Fanuc KAREL source: KS00006.KL

PROGRAM KS00006
%NOLOCKGROUP
TYPE
  REC_T = STRUCTURE
    VALUE: INTEGER
    FLAG: BOOLEAN
  ENDSTRUCTURE
VAR
  A: REC_T
  B: REC_T
  FLAG: BOOLEAN
  N: INTEGER
  STATUS: INTEGER
  PN: STRING[80]
  VN: STRING[80]
BEGIN
  PN = ''
  VN = 'A'
  GET_VAR(N, PN, VN, A, STATUS)
END KS00006
